(* IEC 61131-3 sources: PLC-Static-Analysis/modules/plc-rules/src/test/resources/PLCA-S002, 2 files *)

(* ---- compliant.st ---- *)
VAR_GLOBAL
    GVL_HMI_rSetpoint : REAL;
    GVL_HMI_bRun : BOOL;
    GVL_HMI_nSlot : INT;
    gbFault : BOOL;
    gnInternal : INT;
END_VAR

PROGRAM P_Safe
VAR
    qrOut AT %QD8 : REAL;
    qxRun AT %QX1.0 : BOOL;
    qnOut AT %QW12 : INT;
    arTable : ARRAY[0..9] OF INT;
    n : INT;
END_VAR
qrOut := LIMIT(0.0, GVL_HMI_rSetpoint, 100.0);
qxRun := GVL_HMI_bRun AND NOT gbFault;
qnOut := gnInternal;
IF GVL_HMI_nSlot >= 0 AND GVL_HMI_nSlot <= 9 THEN
    n := arTable[GVL_HMI_nSlot];
END_IF
gnInternal := n;
END_PROGRAM

(* ---- noncompliant.st ---- *)
VAR_GLOBAL
    GVL_HMI_rSpeed : REAL;
    GVL_HMI_bStart : BOOL;
    GVL_HMI_nIndex : INT;
    {attribute 'OPC.UA.DA' := '1'}
    gnRemoteValue : INT;
END_VAR

PROGRAM P_Out
VAR
    qrSpeed AT %QD4 : REAL;
    qxPump AT %QX0.0 : BOOL;
    qxValve AT %QX0.1 : BOOL;
    qnValue AT %QW8 : INT;
    arTable : ARRAY[0..9] OF INT;
    n : INT;
END_VAR
qrSpeed := GVL_HMI_rSpeed * 10.0; // PLCA-S002
qxPump := GVL_HMI_bStart; // PLCA-S002
IF GVL_HMI_bStart THEN
    qxValve := TRUE; // PLCA-S002
END_IF
qnValue := gnRemoteValue; // PLCA-S002
n := arTable[GVL_HMI_nIndex]; // PLCA-S002
END_PROGRAM
